(* IEC 61131-3 sources: STAR-PLC-Agent/results/raw/codex_matrix_resume_20261114/codex_deepseek/SELF005/functional/attempt_0001, 1 file *)

(* ---- test_program.st ---- *)
PROGRAM PLC_PRG
VAR
 BenchStep : UDINT := 0;
 BenchCalls : UDINT := 0;
 BenchDone : BOOL := FALSE;
 BenchUut0 : FB_Task;
 BenchUut1 : FB_Task;
 BenchUut2 : FB_Task;
 BenchUut3 : FB_Task;
 BenchUut4 : FB_Task;
 BenchUut5 : FB_Task;
 BenchUut6 : FB_Task;
 TraceIn_Enable : ARRAY[0..65] OF BOOL;
 TraceIn_Tick : ARRAY[0..65] OF BOOL;
 TraceOut_Red : ARRAY[0..65] OF BOOL;
 TraceOut_Green : ARRAY[0..65] OF BOOL;
 TraceOut_Amber : ARRAY[0..65] OF BOOL;
 TraceOut_Phase : ARRAY[0..65] OF USINT;
END_VAR

IF NOT BenchDone THEN
 CASE BenchStep OF
 0:
   BenchUut0.Enable := TRUE;
   BenchUut0.Tick := TRUE;
   TraceIn_Enable[0] := BenchUut0.Enable;
   TraceIn_Tick[0] := BenchUut0.Tick;
   BenchUut0();
   TraceOut_Red[0] := BenchUut0.Red;
   TraceOut_Green[0] := BenchUut0.Green;
   TraceOut_Amber[0] := BenchUut0.Amber;
   TraceOut_Phase[0] := BenchUut0.Phase;
   BenchCalls := BenchCalls + 1;
 1:
   BenchUut0.Enable := TRUE;
   BenchUut0.Tick := FALSE;
   TraceIn_Enable[1] := BenchUut0.Enable;
   TraceIn_Tick[1] := BenchUut0.Tick;
   BenchUut0();
   TraceOut_Red[1] := BenchUut0.Red;
   TraceOut_Green[1] := BenchUut0.Green;
   TraceOut_Amber[1] := BenchUut0.Amber;
   TraceOut_Phase[1] := BenchUut0.Phase;
   BenchCalls := BenchCalls + 1;
 2:
   BenchUut0.Enable := TRUE;
   BenchUut0.Tick := TRUE;
   TraceIn_Enable[2] := BenchUut0.Enable;
   TraceIn_Tick[2] := BenchUut0.Tick;
   BenchUut0();
   TraceOut_Red[2] := BenchUut0.Red;
   TraceOut_Green[2] := BenchUut0.Green;
   TraceOut_Amber[2] := BenchUut0.Amber;
   TraceOut_Phase[2] := BenchUut0.Phase;
   BenchCalls := BenchCalls + 1;
 3:
   BenchUut0.Enable := TRUE;
   BenchUut0.Tick := TRUE;
   TraceIn_Enable[3] := BenchUut0.Enable;
   TraceIn_Tick[3] := BenchUut0.Tick;
   BenchUut0();
   TraceOut_Red[3] := BenchUut0.Red;
   TraceOut_Green[3] := BenchUut0.Green;
   TraceOut_Amber[3] := BenchUut0.Amber;
   TraceOut_Phase[3] := BenchUut0.Phase;
   BenchCalls := BenchCalls + 1;
 4:
   BenchUut0.Enable := TRUE;
   BenchUut0.Tick := TRUE;
   TraceIn_Enable[4] := BenchUut0.Enable;
   TraceIn_Tick[4] := BenchUut0.Tick;
   BenchUut0();
   TraceOut_Red[4] := BenchUut0.Red;
   TraceOut_Green[4] := BenchUut0.Green;
   TraceOut_Amber[4] := BenchUut0.Amber;
   TraceOut_Phase[4] := BenchUut0.Phase;
   BenchCalls := BenchCalls + 1;
 5:
   BenchUut0.Enable := TRUE;
   BenchUut0.Tick := TRUE;
   TraceIn_Enable[5] := BenchUut0.Enable;
   TraceIn_Tick[5] := BenchUut0.Tick;
   BenchUut0();
   TraceOut_Red[5] := BenchUut0.Red;
   TraceOut_Green[5] := BenchUut0.Green;
   TraceOut_Amber[5] := BenchUut0.Amber;
   TraceOut_Phase[5] := BenchUut0.Phase;
   BenchCalls := BenchCalls + 1;
 6:
   BenchUut0.Enable := TRUE;
   BenchUut0.Tick := TRUE;
   TraceIn_Enable[6] := BenchUut0.Enable;
   TraceIn_Tick[6] := BenchUut0.Tick;
   BenchUut0();
   TraceOut_Red[6] := BenchUut0.Red;
   TraceOut_Green[6] := BenchUut0.Green;
   TraceOut_Amber[6] := BenchUut0.Amber;
   TraceOut_Phase[6] := BenchUut0.Phase;
   BenchCalls := BenchCalls + 1;
 7:
   BenchUut1.Enable := TRUE;
   BenchUut1.Tick := TRUE;
   TraceIn_Enable[7] := BenchUut1.Enable;
   TraceIn_Tick[7] := BenchUut1.Tick;
   BenchUut1();
   TraceOut_Red[7] := BenchUut1.Red;
   TraceOut_Green[7] := BenchUut1.Green;
   TraceOut_Amber[7] := BenchUut1.Amber;
   TraceOut_Phase[7] := BenchUut1.Phase;
   BenchCalls := BenchCalls + 1;
 8:
   BenchUut1.Enable := TRUE;
   BenchUut1.Tick := TRUE;
   TraceIn_Enable[8] := BenchUut1.Enable;
   TraceIn_Tick[8] := BenchUut1.Tick;
   BenchUut1();
   TraceOut_Red[8] := BenchUut1.Red;
   TraceOut_Green[8] := BenchUut1.Green;
   TraceOut_Amber[8] := BenchUut1.Amber;
   TraceOut_Phase[8] := BenchUut1.Phase;
   BenchCalls := BenchCalls + 1;
 9:
   BenchUut1.Enable := FALSE;
   BenchUut1.Tick := TRUE;
   TraceIn_Enable[9] := BenchUut1.Enable;
   TraceIn_Tick[9] := BenchUut1.Tick;
   BenchUut1();
   TraceOut_Red[9] := BenchUut1.Red;
   TraceOut_Green[9] := BenchUut1.Green;
   TraceOut_Amber[9] := BenchUut1.Amber;
   TraceOut_Phase[9] := BenchUut1.Phase;
   BenchCalls := BenchCalls + 1;
 10:
   BenchUut1.Enable := TRUE;
   BenchUut1.Tick := TRUE;
   TraceIn_Enable[10] := BenchUut1.Enable;
   TraceIn_Tick[10] := BenchUut1.Tick;
   BenchUut1();
   TraceOut_Red[10] := BenchUut1.Red;
   TraceOut_Green[10] := BenchUut1.Green;
   TraceOut_Amber[10] := BenchUut1.Amber;
   TraceOut_Phase[10] := BenchUut1.Phase;
   BenchCalls := BenchCalls + 1;
 11:
   BenchUut1.Enable := TRUE;
   BenchUut1.Tick := TRUE;
   TraceIn_Enable[11] := BenchUut1.Enable;
   TraceIn_Tick[11] := BenchUut1.Tick;
   BenchUut1();
   TraceOut_Red[11] := BenchUut1.Red;
   TraceOut_Green[11] := BenchUut1.Green;
   TraceOut_Amber[11] := BenchUut1.Amber;
   TraceOut_Phase[11] := BenchUut1.Phase;
   BenchCalls := BenchCalls + 1;
 12:
   BenchUut2.Enable := TRUE;
   BenchUut2.Tick := TRUE;
   TraceIn_Enable[12] := BenchUut2.Enable;
   TraceIn_Tick[12] := BenchUut2.Tick;
   BenchUut2();
   TraceOut_Red[12] := BenchUut2.Red;
   TraceOut_Green[12] := BenchUut2.Green;
   TraceOut_Amber[12] := BenchUut2.Amber;
   TraceOut_Phase[12] := BenchUut2.Phase;
   BenchCalls := BenchCalls + 1;
 13:
   BenchUut2.Enable := FALSE;
   BenchUut2.Tick := TRUE;
   TraceIn_Enable[13] := BenchUut2.Enable;
   TraceIn_Tick[13] := BenchUut2.Tick;
   BenchUut2();
   TraceOut_Red[13] := BenchUut2.Red;
   TraceOut_Green[13] := BenchUut2.Green;
   TraceOut_Amber[13] := BenchUut2.Amber;
   TraceOut_Phase[13] := BenchUut2.Phase;
   BenchCalls := BenchCalls + 1;
 14:
   BenchUut2.Enable := TRUE;
   BenchUut2.Tick := TRUE;
   TraceIn_Enable[14] := BenchUut2.Enable;
   TraceIn_Tick[14] := BenchUut2.Tick;
   BenchUut2();
   TraceOut_Red[14] := BenchUut2.Red;
   TraceOut_Green[14] := BenchUut2.Green;
   TraceOut_Amber[14] := BenchUut2.Amber;
   TraceOut_Phase[14] := BenchUut2.Phase;
   BenchCalls := BenchCalls + 1;
 15:
   BenchUut2.Enable := TRUE;
   BenchUut2.Tick := TRUE;
   TraceIn_Enable[15] := BenchUut2.Enable;
   TraceIn_Tick[15] := BenchUut2.Tick;
   BenchUut2();
   TraceOut_Red[15] := BenchUut2.Red;
   TraceOut_Green[15] := BenchUut2.Green;
   TraceOut_Amber[15] := BenchUut2.Amber;
   TraceOut_Phase[15] := BenchUut2.Phase;
   BenchCalls := BenchCalls + 1;
 16:
   BenchUut2.Enable := TRUE;
   BenchUut2.Tick := FALSE;
   TraceIn_Enable[16] := BenchUut2.Enable;
   TraceIn_Tick[16] := BenchUut2.Tick;
   BenchUut2();
   TraceOut_Red[16] := BenchUut2.Red;
   TraceOut_Green[16] := BenchUut2.Green;
   TraceOut_Amber[16] := BenchUut2.Amber;
   TraceOut_Phase[16] := BenchUut2.Phase;
   BenchCalls := BenchCalls + 1;
 17:
   BenchUut2.Enable := TRUE;
   BenchUut2.Tick := TRUE;
   TraceIn_Enable[17] := BenchUut2.Enable;
   TraceIn_Tick[17] := BenchUut2.Tick;
   BenchUut2();
   TraceOut_Red[17] := BenchUut2.Red;
   TraceOut_Green[17] := BenchUut2.Green;
   TraceOut_Amber[17] := BenchUut2.Amber;
   TraceOut_Phase[17] := BenchUut2.Phase;
   BenchCalls := BenchCalls + 1;
 18:
   BenchUut2.Enable := TRUE;
   BenchUut2.Tick := TRUE;
   TraceIn_Enable[18] := BenchUut2.Enable;
   TraceIn_Tick[18] := BenchUut2.Tick;
   BenchUut2();
   TraceOut_Red[18] := BenchUut2.Red;
   TraceOut_Green[18] := BenchUut2.Green;
   TraceOut_Amber[18] := BenchUut2.Amber;
   TraceOut_Phase[18] := BenchUut2.Phase;
   BenchCalls := BenchCalls + 1;
 19:
   BenchUut2.Enable := TRUE;
   BenchUut2.Tick := FALSE;
   TraceIn_Enable[19] := BenchUut2.Enable;
   TraceIn_Tick[19] := BenchUut2.Tick;
   BenchUut2();
   TraceOut_Red[19] := BenchUut2.Red;
   TraceOut_Green[19] := BenchUut2.Green;
   TraceOut_Amber[19] := BenchUut2.Amber;
   TraceOut_Phase[19] := BenchUut2.Phase;
   BenchCalls := BenchCalls + 1;
 20:
   BenchUut2.Enable := TRUE;
   BenchUut2.Tick := TRUE;
   TraceIn_Enable[20] := BenchUut2.Enable;
   TraceIn_Tick[20] := BenchUut2.Tick;
   BenchUut2();
   TraceOut_Red[20] := BenchUut2.Red;
   TraceOut_Green[20] := BenchUut2.Green;
   TraceOut_Amber[20] := BenchUut2.Amber;
   TraceOut_Phase[20] := BenchUut2.Phase;
   BenchCalls := BenchCalls + 1;
 21:
   BenchUut2.Enable := TRUE;
   BenchUut2.Tick := TRUE;
   TraceIn_Enable[21] := BenchUut2.Enable;
   TraceIn_Tick[21] := BenchUut2.Tick;
   BenchUut2();
   TraceOut_Red[21] := BenchUut2.Red;
   TraceOut_Green[21] := BenchUut2.Green;
   TraceOut_Amber[21] := BenchUut2.Amber;
   TraceOut_Phase[21] := BenchUut2.Phase;
   BenchCalls := BenchCalls + 1;
 22:
   BenchUut3.Enable := TRUE;
   BenchUut3.Tick := TRUE;
   TraceIn_Enable[22] := BenchUut3.Enable;
   TraceIn_Tick[22] := BenchUut3.Tick;
   BenchUut3();
   TraceOut_Red[22] := BenchUut3.Red;
   TraceOut_Green[22] := BenchUut3.Green;
   TraceOut_Amber[22] := BenchUut3.Amber;
   TraceOut_Phase[22] := BenchUut3.Phase;
   BenchCalls := BenchCalls + 1;
 23:
   BenchUut3.Enable := TRUE;
   BenchUut3.Tick := FALSE;
   TraceIn_Enable[23] := BenchUut3.Enable;
   TraceIn_Tick[23] := BenchUut3.Tick;
   BenchUut3();
   TraceOut_Red[23] := BenchUut3.Red;
   TraceOut_Green[23] := BenchUut3.Green;
   TraceOut_Amber[23] := BenchUut3.Amber;
   TraceOut_Phase[23] := BenchUut3.Phase;
   BenchCalls := BenchCalls + 1;
 24:
   BenchUut3.Enable := TRUE;
   BenchUut3.Tick := TRUE;
   TraceIn_Enable[24] := BenchUut3.Enable;
   TraceIn_Tick[24] := BenchUut3.Tick;
   BenchUut3();
   TraceOut_Red[24] := BenchUut3.Red;
   TraceOut_Green[24] := BenchUut3.Green;
   TraceOut_Amber[24] := BenchUut3.Amber;
   TraceOut_Phase[24] := BenchUut3.Phase;
   BenchCalls := BenchCalls + 1;
 25:
   BenchUut3.Enable := TRUE;
   BenchUut3.Tick := FALSE;
   TraceIn_Enable[25] := BenchUut3.Enable;
   TraceIn_Tick[25] := BenchUut3.Tick;
   BenchUut3();
   TraceOut_Red[25] := BenchUut3.Red;
   TraceOut_Green[25] := BenchUut3.Green;
   TraceOut_Amber[25] := BenchUut3.Amber;
   TraceOut_Phase[25] := BenchUut3.Phase;
   BenchCalls := BenchCalls + 1;
 26:
   BenchUut4.Enable := TRUE;
   BenchUut4.Tick := TRUE;
   TraceIn_Enable[26] := BenchUut4.Enable;
   TraceIn_Tick[26] := BenchUut4.Tick;
   BenchUut4();
   TraceOut_Red[26] := BenchUut4.Red;
   TraceOut_Green[26] := BenchUut4.Green;
   TraceOut_Amber[26] := BenchUut4.Amber;
   TraceOut_Phase[26] := BenchUut4.Phase;
   BenchCalls := BenchCalls + 1;
 27:
   BenchUut4.Enable := TRUE;
   BenchUut4.Tick := FALSE;
   TraceIn_Enable[27] := BenchUut4.Enable;
   TraceIn_Tick[27] := BenchUut4.Tick;
   BenchUut4();
   TraceOut_Red[27] := BenchUut4.Red;
   TraceOut_Green[27] := BenchUut4.Green;
   TraceOut_Amber[27] := BenchUut4.Amber;
   TraceOut_Phase[27] := BenchUut4.Phase;
   BenchCalls := BenchCalls + 1;
 28:
   BenchUut4.Enable := TRUE;
   BenchUut4.Tick := TRUE;
   TraceIn_Enable[28] := BenchUut4.Enable;
   TraceIn_Tick[28] := BenchUut4.Tick;
   BenchUut4();
   TraceOut_Red[28] := BenchUut4.Red;
   TraceOut_Green[28] := BenchUut4.Green;
   TraceOut_Amber[28] := BenchUut4.Amber;
   TraceOut_Phase[28] := BenchUut4.Phase;
   BenchCalls := BenchCalls + 1;
 29:
   BenchUut4.Enable := TRUE;
   BenchUut4.Tick := FALSE;
   TraceIn_Enable[29] := BenchUut4.Enable;
   TraceIn_Tick[29] := BenchUut4.Tick;
   BenchUut4();
   TraceOut_Red[29] := BenchUut4.Red;
   TraceOut_Green[29] := BenchUut4.Green;
   TraceOut_Amber[29] := BenchUut4.Amber;
   TraceOut_Phase[29] := BenchUut4.Phase;
   BenchCalls := BenchCalls + 1;
 30:
   BenchUut4.Enable := TRUE;
   BenchUut4.Tick := TRUE;
   TraceIn_Enable[30] := BenchUut4.Enable;
   TraceIn_Tick[30] := BenchUut4.Tick;
   BenchUut4();
   TraceOut_Red[30] := BenchUut4.Red;
   TraceOut_Green[30] := BenchUut4.Green;
   TraceOut_Amber[30] := BenchUut4.Amber;
   TraceOut_Phase[30] := BenchUut4.Phase;
   BenchCalls := BenchCalls + 1;
 31:
   BenchUut4.Enable := TRUE;
   BenchUut4.Tick := FALSE;
   TraceIn_Enable[31] := BenchUut4.Enable;
   TraceIn_Tick[31] := BenchUut4.Tick;
   BenchUut4();
   TraceOut_Red[31] := BenchUut4.Red;
   TraceOut_Green[31] := BenchUut4.Green;
   TraceOut_Amber[31] := BenchUut4.Amber;
   TraceOut_Phase[31] := BenchUut4.Phase;
   BenchCalls := BenchCalls + 1;
 32:
   BenchUut4.Enable := TRUE;
   BenchUut4.Tick := TRUE;
   TraceIn_Enable[32] := BenchUut4.Enable;
   TraceIn_Tick[32] := BenchUut4.Tick;
   BenchUut4();
   TraceOut_Red[32] := BenchUut4.Red;
   TraceOut_Green[32] := BenchUut4.Green;
   TraceOut_Amber[32] := BenchUut4.Amber;
   TraceOut_Phase[32] := BenchUut4.Phase;
   BenchCalls := BenchCalls + 1;
 33:
   BenchUut4.Enable := TRUE;
   BenchUut4.Tick := FALSE;
   TraceIn_Enable[33] := BenchUut4.Enable;
   TraceIn_Tick[33] := BenchUut4.Tick;
   BenchUut4();
   TraceOut_Red[33] := BenchUut4.Red;
   TraceOut_Green[33] := BenchUut4.Green;
   TraceOut_Amber[33] := BenchUut4.Amber;
   TraceOut_Phase[33] := BenchUut4.Phase;
   BenchCalls := BenchCalls + 1;
 34:
   BenchUut4.Enable := TRUE;
   BenchUut4.Tick := TRUE;
   TraceIn_Enable[34] := BenchUut4.Enable;
   TraceIn_Tick[34] := BenchUut4.Tick;
   BenchUut4();
   TraceOut_Red[34] := BenchUut4.Red;
   TraceOut_Green[34] := BenchUut4.Green;
   TraceOut_Amber[34] := BenchUut4.Amber;
   TraceOut_Phase[34] := BenchUut4.Phase;
   BenchCalls := BenchCalls + 1;
 35:
   BenchUut4.Enable := TRUE;
   BenchUut4.Tick := FALSE;
   TraceIn_Enable[35] := BenchUut4.Enable;
   TraceIn_Tick[35] := BenchUut4.Tick;
   BenchUut4();
   TraceOut_Red[35] := BenchUut4.Red;
   TraceOut_Green[35] := BenchUut4.Green;
   TraceOut_Amber[35] := BenchUut4.Amber;
   TraceOut_Phase[35] := BenchUut4.Phase;
   BenchCalls := BenchCalls + 1;
 36:
   BenchUut4.Enable := TRUE;
   BenchUut4.Tick := TRUE;
   TraceIn_Enable[36] := BenchUut4.Enable;
   TraceIn_Tick[36] := BenchUut4.Tick;
   BenchUut4();
   TraceOut_Red[36] := BenchUut4.Red;
   TraceOut_Green[36] := BenchUut4.Green;
   TraceOut_Amber[36] := BenchUut4.Amber;
   TraceOut_Phase[36] := BenchUut4.Phase;
   BenchCalls := BenchCalls + 1;
 37:
   BenchUut4.Enable := TRUE;
   BenchUut4.Tick := TRUE;
   TraceIn_Enable[37] := BenchUut4.Enable;
   TraceIn_Tick[37] := BenchUut4.Tick;
   BenchUut4();
   TraceOut_Red[37] := BenchUut4.Red;
   TraceOut_Green[37] := BenchUut4.Green;
   TraceOut_Amber[37] := BenchUut4.Amber;
   TraceOut_Phase[37] := BenchUut4.Phase;
   BenchCalls := BenchCalls + 1;
 38:
   BenchUut4.Enable := TRUE;
   BenchUut4.Tick := FALSE;
   TraceIn_Enable[38] := BenchUut4.Enable;
   TraceIn_Tick[38] := BenchUut4.Tick;
   BenchUut4();
   TraceOut_Red[38] := BenchUut4.Red;
   TraceOut_Green[38] := BenchUut4.Green;
   TraceOut_Amber[38] := BenchUut4.Amber;
   TraceOut_Phase[38] := BenchUut4.Phase;
   BenchCalls := BenchCalls + 1;
 39:
   BenchUut4.Enable := TRUE;
   BenchUut4.Tick := TRUE;
   TraceIn_Enable[39] := BenchUut4.Enable;
   TraceIn_Tick[39] := BenchUut4.Tick;
   BenchUut4();
   TraceOut_Red[39] := BenchUut4.Red;
   TraceOut_Green[39] := BenchUut4.Green;
   TraceOut_Amber[39] := BenchUut4.Amber;
   TraceOut_Phase[39] := BenchUut4.Phase;
   BenchCalls := BenchCalls + 1;
 40:
   BenchUut4.Enable := TRUE;
   BenchUut4.Tick := FALSE;
   TraceIn_Enable[40] := BenchUut4.Enable;
   TraceIn_Tick[40] := BenchUut4.Tick;
   BenchUut4();
   TraceOut_Red[40] := BenchUut4.Red;
   TraceOut_Green[40] := BenchUut4.Green;
   TraceOut_Amber[40] := BenchUut4.Amber;
   TraceOut_Phase[40] := BenchUut4.Phase;
   BenchCalls := BenchCalls + 1;
 41:
   BenchUut4.Enable := TRUE;
   BenchUut4.Tick := TRUE;
   TraceIn_Enable[41] := BenchUut4.Enable;
   TraceIn_Tick[41] := BenchUut4.Tick;
   BenchUut4();
   TraceOut_Red[41] := BenchUut4.Red;
   TraceOut_Green[41] := BenchUut4.Green;
   TraceOut_Amber[41] := BenchUut4.Amber;
   TraceOut_Phase[41] := BenchUut4.Phase;
   BenchCalls := BenchCalls + 1;
 42:
   BenchUut4.Enable := TRUE;
   BenchUut4.Tick := FALSE;
   TraceIn_Enable[42] := BenchUut4.Enable;
   TraceIn_Tick[42] := BenchUut4.Tick;
   BenchUut4();
   TraceOut_Red[42] := BenchUut4.Red;
   TraceOut_Green[42] := BenchUut4.Green;
   TraceOut_Amber[42] := BenchUut4.Amber;
   TraceOut_Phase[42] := BenchUut4.Phase;
   BenchCalls := BenchCalls + 1;
 43:
   BenchUut4.Enable := TRUE;
   BenchUut4.Tick := TRUE;
   TraceIn_Enable[43] := BenchUut4.Enable;
   TraceIn_Tick[43] := BenchUut4.Tick;
   BenchUut4();
   TraceOut_Red[43] := BenchUut4.Red;
   TraceOut_Green[43] := BenchUut4.Green;
   TraceOut_Amber[43] := BenchUut4.Amber;
   TraceOut_Phase[43] := BenchUut4.Phase;
   BenchCalls := BenchCalls + 1;
 44:
   BenchUut4.Enable := TRUE;
   BenchUut4.Tick := FALSE;
   TraceIn_Enable[44] := BenchUut4.Enable;
   TraceIn_Tick[44] := BenchUut4.Tick;
   BenchUut4();
   TraceOut_Red[44] := BenchUut4.Red;
   TraceOut_Green[44] := BenchUut4.Green;
   TraceOut_Amber[44] := BenchUut4.Amber;
   TraceOut_Phase[44] := BenchUut4.Phase;
   BenchCalls := BenchCalls + 1;
 45:
   BenchUut4.Enable := TRUE;
   BenchUut4.Tick := TRUE;
   TraceIn_Enable[45] := BenchUut4.Enable;
   TraceIn_Tick[45] := BenchUut4.Tick;
   BenchUut4();
   TraceOut_Red[45] := BenchUut4.Red;
   TraceOut_Green[45] := BenchUut4.Green;
   TraceOut_Amber[45] := BenchUut4.Amber;
   TraceOut_Phase[45] := BenchUut4.Phase;
   BenchCalls := BenchCalls + 1;
 46:
   BenchUut4.Enable := TRUE;
   BenchUut4.Tick := FALSE;
   TraceIn_Enable[46] := BenchUut4.Enable;
   TraceIn_Tick[46] := BenchUut4.Tick;
   BenchUut4();
   TraceOut_Red[46] := BenchUut4.Red;
   TraceOut_Green[46] := BenchUut4.Green;
   TraceOut_Amber[46] := BenchUut4.Amber;
   TraceOut_Phase[46] := BenchUut4.Phase;
   BenchCalls := BenchCalls + 1;
 47:
   BenchUut4.Enable := TRUE;
   BenchUut4.Tick := TRUE;
   TraceIn_Enable[47] := BenchUut4.Enable;
   TraceIn_Tick[47] := BenchUut4.Tick;
   BenchUut4();
   TraceOut_Red[47] := BenchUut4.Red;
   TraceOut_Green[47] := BenchUut4.Green;
   TraceOut_Amber[47] := BenchUut4.Amber;
   TraceOut_Phase[47] := BenchUut4.Phase;
   BenchCalls := BenchCalls + 1;
 48:
   BenchUut5.Enable := TRUE;
   BenchUut5.Tick := TRUE;
   TraceIn_Enable[48] := BenchUut5.Enable;
   TraceIn_Tick[48] := BenchUut5.Tick;
   BenchUut5();
   TraceOut_Red[48] := BenchUut5.Red;
   TraceOut_Green[48] := BenchUut5.Green;
   TraceOut_Amber[48] := BenchUut5.Amber;
   TraceOut_Phase[48] := BenchUut5.Phase;
   BenchCalls := BenchCalls + 1;
 49:
   BenchUut5.Enable := TRUE;
   BenchUut5.Tick := FALSE;
   TraceIn_Enable[49] := BenchUut5.Enable;
   TraceIn_Tick[49] := BenchUut5.Tick;
   BenchUut5();
   TraceOut_Red[49] := BenchUut5.Red;
   TraceOut_Green[49] := BenchUut5.Green;
   TraceOut_Amber[49] := BenchUut5.Amber;
   TraceOut_Phase[49] := BenchUut5.Phase;
   BenchCalls := BenchCalls + 1;
 50:
   BenchUut5.Enable := TRUE;
   BenchUut5.Tick := TRUE;
   TraceIn_Enable[50] := BenchUut5.Enable;
   TraceIn_Tick[50] := BenchUut5.Tick;
   BenchUut5();
   TraceOut_Red[50] := BenchUut5.Red;
   TraceOut_Green[50] := BenchUut5.Green;
   TraceOut_Amber[50] := BenchUut5.Amber;
   TraceOut_Phase[50] := BenchUut5.Phase;
   BenchCalls := BenchCalls + 1;
 51:
   BenchUut5.Enable := TRUE;
   BenchUut5.Tick := TRUE;
   TraceIn_Enable[51] := BenchUut5.Enable;
   TraceIn_Tick[51] := BenchUut5.Tick;
   BenchUut5();
   TraceOut_Red[51] := BenchUut5.Red;
   TraceOut_Green[51] := BenchUut5.Green;
   TraceOut_Amber[51] := BenchUut5.Amber;
   TraceOut_Phase[51] := BenchUut5.Phase;
   BenchCalls := BenchCalls + 1;
 52:
   BenchUut5.Enable := TRUE;
   BenchUut5.Tick := TRUE;
   TraceIn_Enable[52] := BenchUut5.Enable;
   TraceIn_Tick[52] := BenchUut5.Tick;
   BenchUut5();
   TraceOut_Red[52] := BenchUut5.Red;
   TraceOut_Green[52] := BenchUut5.Green;
   TraceOut_Amber[52] := BenchUut5.Amber;
   TraceOut_Phase[52] := BenchUut5.Phase;
   BenchCalls := BenchCalls + 1;
 53:
   BenchUut5.Enable := TRUE;
   BenchUut5.Tick := TRUE;
   TraceIn_Enable[53] := BenchUut5.Enable;
   TraceIn_Tick[53] := BenchUut5.Tick;
   BenchUut5();
   TraceOut_Red[53] := BenchUut5.Red;
   TraceOut_Green[53] := BenchUut5.Green;
   TraceOut_Amber[53] := BenchUut5.Amber;
   TraceOut_Phase[53] := BenchUut5.Phase;
   BenchCalls := BenchCalls + 1;
 54:
   BenchUut5.Enable := TRUE;
   BenchUut5.Tick := TRUE;
   TraceIn_Enable[54] := BenchUut5.Enable;
   TraceIn_Tick[54] := BenchUut5.Tick;
   BenchUut5();
   TraceOut_Red[54] := BenchUut5.Red;
   TraceOut_Green[54] := BenchUut5.Green;
   TraceOut_Amber[54] := BenchUut5.Amber;
   TraceOut_Phase[54] := BenchUut5.Phase;
   BenchCalls := BenchCalls + 1;
 55:
   BenchUut5.Enable := FALSE;
   BenchUut5.Tick := TRUE;
   TraceIn_Enable[55] := BenchUut5.Enable;
   TraceIn_Tick[55] := BenchUut5.Tick;
   BenchUut5();
   TraceOut_Red[55] := BenchUut5.Red;
   TraceOut_Green[55] := BenchUut5.Green;
   TraceOut_Amber[55] := BenchUut5.Amber;
   TraceOut_Phase[55] := BenchUut5.Phase;
   BenchCalls := BenchCalls + 1;
 56:
   BenchUut5.Enable := FALSE;
   BenchUut5.Tick := TRUE;
   TraceIn_Enable[56] := BenchUut5.Enable;
   TraceIn_Tick[56] := BenchUut5.Tick;
   BenchUut5();
   TraceOut_Red[56] := BenchUut5.Red;
   TraceOut_Green[56] := BenchUut5.Green;
   TraceOut_Amber[56] := BenchUut5.Amber;
   TraceOut_Phase[56] := BenchUut5.Phase;
   BenchCalls := BenchCalls + 1;
 57:
   BenchUut6.Enable := TRUE;
   BenchUut6.Tick := TRUE;
   TraceIn_Enable[57] := BenchUut6.Enable;
   TraceIn_Tick[57] := BenchUut6.Tick;
   BenchUut6();
   TraceOut_Red[57] := BenchUut6.Red;
   TraceOut_Green[57] := BenchUut6.Green;
   TraceOut_Amber[57] := BenchUut6.Amber;
   TraceOut_Phase[57] := BenchUut6.Phase;
   BenchCalls := BenchCalls + 1;
 58:
   BenchUut6.Enable := TRUE;
   BenchUut6.Tick := FALSE;
   TraceIn_Enable[58] := BenchUut6.Enable;
   TraceIn_Tick[58] := BenchUut6.Tick;
   BenchUut6();
   TraceOut_Red[58] := BenchUut6.Red;
   TraceOut_Green[58] := BenchUut6.Green;
   TraceOut_Amber[58] := BenchUut6.Amber;
   TraceOut_Phase[58] := BenchUut6.Phase;
   BenchCalls := BenchCalls + 1;
 59:
   BenchUut6.Enable := TRUE;
   BenchUut6.Tick := TRUE;
   TraceIn_Enable[59] := BenchUut6.Enable;
   TraceIn_Tick[59] := BenchUut6.Tick;
   BenchUut6();
   TraceOut_Red[59] := BenchUut6.Red;
   TraceOut_Green[59] := BenchUut6.Green;
   TraceOut_Amber[59] := BenchUut6.Amber;
   TraceOut_Phase[59] := BenchUut6.Phase;
   BenchCalls := BenchCalls + 1;
 60:
   BenchUut6.Enable := TRUE;
   BenchUut6.Tick := TRUE;
   TraceIn_Enable[60] := BenchUut6.Enable;
   TraceIn_Tick[60] := BenchUut6.Tick;
   BenchUut6();
   TraceOut_Red[60] := BenchUut6.Red;
   TraceOut_Green[60] := BenchUut6.Green;
   TraceOut_Amber[60] := BenchUut6.Amber;
   TraceOut_Phase[60] := BenchUut6.Phase;
   BenchCalls := BenchCalls + 1;
 61:
   BenchUut6.Enable := TRUE;
   BenchUut6.Tick := TRUE;
   TraceIn_Enable[61] := BenchUut6.Enable;
   TraceIn_Tick[61] := BenchUut6.Tick;
   BenchUut6();
   TraceOut_Red[61] := BenchUut6.Red;
   TraceOut_Green[61] := BenchUut6.Green;
   TraceOut_Amber[61] := BenchUut6.Amber;
   TraceOut_Phase[61] := BenchUut6.Phase;
   BenchCalls := BenchCalls + 1;
 62:
   BenchUut6.Enable := TRUE;
   BenchUut6.Tick := TRUE;
   TraceIn_Enable[62] := BenchUut6.Enable;
   TraceIn_Tick[62] := BenchUut6.Tick;
   BenchUut6();
   TraceOut_Red[62] := BenchUut6.Red;
   TraceOut_Green[62] := BenchUut6.Green;
   TraceOut_Amber[62] := BenchUut6.Amber;
   TraceOut_Phase[62] := BenchUut6.Phase;
   BenchCalls := BenchCalls + 1;
 63:
   BenchUut6.Enable := TRUE;
   BenchUut6.Tick := TRUE;
   TraceIn_Enable[63] := BenchUut6.Enable;
   TraceIn_Tick[63] := BenchUut6.Tick;
   BenchUut6();
   TraceOut_Red[63] := BenchUut6.Red;
   TraceOut_Green[63] := BenchUut6.Green;
   TraceOut_Amber[63] := BenchUut6.Amber;
   TraceOut_Phase[63] := BenchUut6.Phase;
   BenchCalls := BenchCalls + 1;
 64:
   BenchUut6.Enable := TRUE;
   BenchUut6.Tick := FALSE;
   TraceIn_Enable[64] := BenchUut6.Enable;
   TraceIn_Tick[64] := BenchUut6.Tick;
   BenchUut6();
   TraceOut_Red[64] := BenchUut6.Red;
   TraceOut_Green[64] := BenchUut6.Green;
   TraceOut_Amber[64] := BenchUut6.Amber;
   TraceOut_Phase[64] := BenchUut6.Phase;
   BenchCalls := BenchCalls + 1;
 65:
   BenchUut6.Enable := TRUE;
   BenchUut6.Tick := FALSE;
   TraceIn_Enable[65] := BenchUut6.Enable;
   TraceIn_Tick[65] := BenchUut6.Tick;
   BenchUut6();
   TraceOut_Red[65] := BenchUut6.Red;
   TraceOut_Green[65] := BenchUut6.Green;
   TraceOut_Amber[65] := BenchUut6.Amber;
   TraceOut_Phase[65] := BenchUut6.Phase;
   BenchCalls := BenchCalls + 1;
 END_CASE;
 BenchStep := BenchStep + 1;
 IF BenchStep >= 66 THEN BenchDone := TRUE; END_IF;
END_IF;
END_PROGRAM
